TYPE E_SlideState :
(
    eSlideOut    := 0,
    eSlideIn     := 1,
    eSlideMoving := 2,
    eSlideError  := 3
) INT;
END_TYPE

(* stored: Version 1.1.0.1, ProductVersion 3.1.4026.18
   DUT E_SlideState: Id {bbf93ea1-6e2a-4304-83a7-82d06f1646ae} *)
